(* IEC 61131-3 sources: Caravan/Archiv/12-04-19/Stations/MachineControl/MachineControl/Network/LseEasyMain, 1 file *)

(* ---- ONE_LseEasyMain_Table.st ---- *)
#define OBJECTS_CONFIG

#include "..\..\Source\Common\hmi_nuc.h"

FUNCTION GLOBAL TAB ONE_LseEasyMain
-1$UINT, 0$UINT,
0$UINT, 0$UINT,

40$UDINT,
TO_UDINT(3253426089), "HmiAsciiBuffer", 0$UINT, 0$UINT, 4$UINT,
TO_UDINT(3735923847), "HmiBaseList", 0$UINT, 0$UINT, 0$UINT,
TO_UDINT(2189921946), "HmiCanSendReceive", 0$UINT, 2$UINT, 1$UINT,
TO_UDINT(3930770040), "HmiChkBitList", 0$UINT, 2$UINT, 1$UINT,
TO_UDINT(845038353), "HmiColorMap", 0$UINT, 0$UINT, 1$UINT,
TO_UDINT(136722037), "HmiComPort", 0$UINT, 15$UINT, 0$UINT,
TO_UDINT(4239410787), "HmiComPortCan", 0$UINT, 14$UINT, 1$UINT,
TO_UDINT(2548286290), "HmiFile", 0$UINT, 4$UINT, 2$UINT,
TO_UDINT(1363967167), "HmiFont35", 0$UINT, 1$UINT, 1$UINT,
TO_UDINT(3893392983), "HmiFontList", 0$UINT, 3$UINT, 1$UINT,
TO_UDINT(3842677476), "HmiFunctionList", 0$UINT, 2$UINT, 1$UINT,
TO_UDINT(3385399892), "HmiFunctionList35", 0$UINT, 3$UINT, 1$UINT,
TO_UDINT(2724513001), "HmiImage35", 0$UINT, 3$UINT, 1$UINT,
TO_UDINT(3242935315), "HmiImageList", 0$UINT, 3$UINT, 1$UINT,
TO_UDINT(896341175), "HmiMapFile", 0$UINT, 0$UINT, 1$UINT,
TO_UDINT(3426238687), "HmiMemCircle", 0$UINT, 0$UINT, 1$UINT,
TO_UDINT(4250916264), "HmiMemImage", 0$UINT, 0$UINT, 1$UINT,
TO_UDINT(568511237), "HmiMemIO", 0$UINT, 0$UINT, 1$UINT,
TO_UDINT(1795655540), "HmiMemLine", 0$UINT, 0$UINT, 1$UINT,
TO_UDINT(2462046095), "HmiMemRectangle", 0$UINT, 0$UINT, 1$UINT,
TO_UDINT(2174260293), "HmiMemText", 0$UINT, 0$UINT, 1$UINT,
TO_UDINT(822070823), "HmiMemZorder", 0$UINT, 0$UINT, 1$UINT,
TO_UDINT(2613567777), "HmiProject35", 0$UINT, 4$UINT, 1$UINT,
TO_UDINT(2305619121), "HmiProjectList", 0$UINT, 1$UINT, 1$UINT,
TO_UDINT(2118014258), "HmiScreen", 0$UINT, 1$UINT, 1$UINT,
TO_UDINT(4172848962), "HmiSetUpList", 0$UINT, 2$UINT, 1$UINT,
TO_UDINT(1107224582), "HmiSetupList35", 0$UINT, 2$UINT, 1$UINT,
TO_UDINT(3851519469), "HmiShemeList", 0$UINT, 3$UINT, 4$UINT,
TO_UDINT(2500045939), "HmiShemeList35", 0$UINT, 3$UINT, 1$UINT,
TO_UDINT(4141094888), "HmiStateBit35", 0$UINT, 4$UINT, 1$UINT,
TO_UDINT(103556616), "HmiStrLib", 0$UINT, 2$UINT, 1$UINT,
TO_UDINT(2809265865), "HmiTextList", 0$UINT, 3$UINT, 1$UINT,
TO_UDINT(2738661249), "HmiTextList35", 0$UINT, 1$UINT, 1$UINT,
TO_UDINT(2548567416), "HmiUniBuffer", 0$UINT, 0$UINT, 10$UINT,
TO_UDINT(2706799507), "HmiUnitList", 0$UINT, 2$UINT, 1$UINT,
TO_UDINT(4154992490), "HmiUtils", 0$UINT, 2$UINT, 1$UINT,
TO_UDINT(1002095878), "HmiVarInfoList", 0$UINT, 1$UINT, 1$UINT,
TO_UDINT(3793961451), "HmiVarList", 0$UINT, 15$UINT, 1$UINT,
TO_UDINT(1599081198), "HmiVarList35", 0$UINT, 4$UINT, 1$UINT,
TO_UDINT(1518191916), "LseEasy", 1$UINT, 26$UINT, 1$UINT,

1$UINT, TO_UDINT(1344493304), "LSEEASY\HMICHKBITLIST\LABEL",
1$UINT, TO_UDINT(787249025), "LSEEASY\HMIFONTLIST\LABEL",
1$UINT, TO_UDINT(2117594790), "LSEEASY\HMIIMAGELIST\LABEL",
1$UINT, TO_UDINT(3002767849), "LSEEASY\HMIVARLIST\LABEL",

1$UINT, TO_UDINT(4084571679), "HMICOMPORTCAN1\CANSEND",

1$UINT, TO_UDINT(4275455085), "LSEEASY\HMICHKBITLIST",

1$UINT, TO_UDINT(846459028), "LSEEASY\HMICOLORMAP",

_NO_ATTR, TO_UDINT(1469804307), "HMICOMPORTCAN1",

1$UINT, TO_UDINT(1873895348), "HMICOMPORTCAN1\_BASE\FILE",
1$UINT, TO_UDINT(4182786947), "LSEEASY\FILE",

1$UINT, TO_UDINT(3760648512), "LSEEASY\HMIFONT35",

1$UINT, TO_UDINT(3896362450), "LSEEASY\HMIFONTLIST",

1$UINT, TO_UDINT(3636446795), "LSEEASY\HMIFUNCTIONLIST",

1$UINT, TO_UDINT(2190187032), "LSEEASY\HMIFUNCTIONLIST35",

1$UINT, TO_UDINT(2413249001), "LSEEASY\HMIIMAGE35",

1$UINT, TO_UDINT(1553538575), "LSEEASY\HMIIMAGELIST",

1$UINT, TO_UDINT(417239479), "LSEEASY\HMIMAPFILE",

1$UINT, TO_UDINT(2012497378), "LSEEASY\HMISCREEN\MEMCIRCLE",

1$UINT, TO_UDINT(975039261), "LSEEASY\HMISCREEN\MEMIMAGE",

1$UINT, TO_UDINT(3016924028), "LSEEASY\HMISCREEN\MEMIO",

1$UINT, TO_UDINT(4270949903), "LSEEASY\HMISCREEN\MEMLINE",

1$UINT, TO_UDINT(1370086185), "LSEEASY\HMISCREEN\MEMRECTANGLE",

1$UINT, TO_UDINT(336500030), "LSEEASY\HMISCREEN\MEMTEXT",

1$UINT, TO_UDINT(2335427354), "LSEEASY\HMISCREEN\MEMZORDER",

1$UINT, TO_UDINT(102087485), "LSEEASY\HMIPROJECT35",

1$UINT, TO_UDINT(3836054740), "LSEEASY\HMIPROJECTLIST",

1$UINT, TO_UDINT(3478444237), "LSEEASY\HMISCREEN",

1$UINT, TO_UDINT(1701496158), "LSEEASY\HMISETUPLIST",

1$UINT, TO_UDINT(741838947), "LSEEASY\HMISETUPLIST35",

1$UINT, TO_UDINT(2459869223), "LSEEASY\HMIFONTSHEMELIST",
1$UINT, TO_UDINT(1282849623), "LSEEASY\HMIIMAGESHEMELIST",
1$UINT, TO_UDINT(3937490271), "LSEEASY\HMITEXTSHEMELIST",
1$UINT, TO_UDINT(3509062318), "LSEEASY\HMIVARLIST\HMIUNITSHEMELIST",

1$UINT, TO_UDINT(4174042134), "LSEEASY\HMISHEMELIST35",

1$UINT, TO_UDINT(3796408829), "LSEEASY\HMISTATEBIT35",

1$UINT, TO_UDINT(1881447452), "LSEEASY\STRINGLIB",

1$UINT, TO_UDINT(2807844172), "LSEEASY\HMITEXTLIST",

1$UINT, TO_UDINT(3080726932), "LSEEASY\HMITEXTLIST35",

1$UINT, TO_UDINT(2308124733), "LSEEASY\HMITEXTLIST\TEXTLIST00",
1$UINT, TO_UDINT(4271112363), "LSEEASY\HMITEXTLIST\TEXTLIST01",
1$UINT, TO_UDINT(1738363153), "LSEEASY\HMITEXTLIST\TEXTLIST02",
1$UINT, TO_UDINT(278552967), "LSEEASY\HMITEXTLIST\TEXTLIST03",
1$UINT, TO_UDINT(2399073316), "LSEEASY\HMITEXTLIST\TEXTLIST04",
1$UINT, TO_UDINT(4193895602), "LSEEASY\HMITEXTLIST\TEXTLIST05",
1$UINT, TO_UDINT(1626379528), "LSEEASY\HMITEXTLIST\TEXTLIST06",
1$UINT, TO_UDINT(402105758), "LSEEASY\HMITEXTLIST\TEXTLIST07",
1$UINT, TO_UDINT(2269689871), "LSEEASY\HMITEXTLIST\TEXTLIST08",
1$UINT, TO_UDINT(4031744153), "LSEEASY\HMITEXTLIST\TEXTLIST09",

1$UINT, TO_UDINT(200861884), "LSEEASY\HMIVARLIST\UNITINFO",

1$UINT, TO_UDINT(2530016337), "LSEEASY\HMIUTILS",

1$UINT, TO_UDINT(3991554070), "LSEEASY\HMIVARLIST\VARINFO",

1$UINT, TO_UDINT(3482371307), "LSEEASY\HMIVARLIST",

1$UINT, TO_UDINT(3263320306), "LSEEASY\HMIVARLIST35",

_NO_ATTR, TO_UDINT(1518191916), "LSEEASY",

//Internal connections
0$UDINT,
52$UDINT,
TO_UDINT(5), "Label", TO_UDINT(0),
TO_UDINT(7), "File", TO_UDINT(8),
TO_UDINT(7), "CanSend", TO_UDINT(4),
TO_UDINT(11), "Label", TO_UDINT(1),
TO_UDINT(15), "Label", TO_UDINT(2),
TO_UDINT(26), "MemRectangle", TO_UDINT(21),
TO_UDINT(26), "MemText", TO_UDINT(22),
TO_UDINT(26), "MemIO", TO_UDINT(19),
TO_UDINT(26), "MemCircle", TO_UDINT(17),
TO_UDINT(26), "MemLine", TO_UDINT(20),
TO_UDINT(26), "MemImage", TO_UDINT(18),
TO_UDINT(26), "MemZorder", TO_UDINT(23),
TO_UDINT(36), "TextList00", TO_UDINT(38),
TO_UDINT(36), "TextList01", TO_UDINT(39),
TO_UDINT(36), "TextList02", TO_UDINT(40),
TO_UDINT(36), "TextList03", TO_UDINT(41),
TO_UDINT(36), "TextList04", TO_UDINT(42),
TO_UDINT(36), "TextList05", TO_UDINT(43),
TO_UDINT(36), "TextList06", TO_UDINT(44),
TO_UDINT(36), "TextList07", TO_UDINT(45),
TO_UDINT(36), "TextList08", TO_UDINT(46),
TO_UDINT(36), "TextList09", TO_UDINT(47),
TO_UDINT(51), "UnitInfo", TO_UDINT(48),
TO_UDINT(51), "Label", TO_UDINT(3),
TO_UDINT(51), "VarInfo", TO_UDINT(50),
TO_UDINT(51), "HmiUnitShemeList", TO_UDINT(32),
TO_UDINT(53), "HmiImageList", TO_UDINT(15),
TO_UDINT(53), "HmiFunctionList", TO_UDINT(12),
TO_UDINT(53), "HmiScreen", TO_UDINT(26),
TO_UDINT(53), "HmiFontList", TO_UDINT(11),
TO_UDINT(53), "HmiVarList", TO_UDINT(51),
TO_UDINT(53), "HmiColorMap", TO_UDINT(6),
TO_UDINT(53), "HmiProjectList", TO_UDINT(25),
TO_UDINT(53), "HmiProject35", TO_UDINT(24),
TO_UDINT(53), "HmiTextList", TO_UDINT(36),
TO_UDINT(53), "HmiVarList35", TO_UDINT(52),
TO_UDINT(53), "HmiFont35", TO_UDINT(10),
TO_UDINT(53), "HmiImage35", TO_UDINT(14),
TO_UDINT(53), "HmiSetUpList", TO_UDINT(27),
TO_UDINT(53), "HmiFunctionList35", TO_UDINT(13),
TO_UDINT(53), "HmiShemeList35", TO_UDINT(33),
TO_UDINT(53), "HmiFontShemeList", TO_UDINT(29),
TO_UDINT(53), "HmiTextShemeList", TO_UDINT(31),
TO_UDINT(53), "HmiImageShemeList", TO_UDINT(30),
TO_UDINT(53), "HmiSetupList35", TO_UDINT(28),
TO_UDINT(53), "StringLib", TO_UDINT(35),
TO_UDINT(53), "File", TO_UDINT(9),
TO_UDINT(53), "HmiUtils", TO_UDINT(49),
TO_UDINT(53), "HmiTextList35", TO_UDINT(37),
TO_UDINT(53), "HmiChkBitList", TO_UDINT(5),
TO_UDINT(53), "HmiStateBit35", TO_UDINT(34),
TO_UDINT(53), "HmiMapFile", TO_UDINT(16),
0$UDINT,
33$UDINT,
TO_UDINT(5), "File", TO_UDINT(9), "ClassSvr",
TO_UDINT(5), "VarList", TO_UDINT(51), "ClassSvr",
TO_UDINT(5), "StringLib", TO_UDINT(35), "ClassSvr",
TO_UDINT(6), "File", TO_UDINT(9), "ClassSvr",
TO_UDINT(11), "File", TO_UDINT(9), "ClassSvr",
TO_UDINT(11), "StringLib", TO_UDINT(35), "ClassSvr",
TO_UDINT(12), "File", TO_UDINT(9), "ClassSvr",
TO_UDINT(13), "HmiVarList", TO_UDINT(51), "ClassSvr",
TO_UDINT(15), "File", TO_UDINT(9), "ClassSvr",
TO_UDINT(15), "StringLib", TO_UDINT(35), "ClassSvr",
TO_UDINT(16), "File", TO_UDINT(9), "ClassSvr",
TO_UDINT(16), "VarList", TO_UDINT(51), "ClassSvr",
TO_UDINT(16), "StateBit", TO_UDINT(34), "ClassSvr",
TO_UDINT(16), "StringLib", TO_UDINT(35), "ClassSvr",
TO_UDINT(25), "File", TO_UDINT(9), "ClassSvr",
TO_UDINT(25), "StringLib", TO_UDINT(35), "ClassSvr",
TO_UDINT(26), "File", TO_UDINT(9), "ClassSvr",
TO_UDINT(27), "File", TO_UDINT(9), "ClassSvr",
TO_UDINT(29), "File", TO_UDINT(9), "ClassSvr",
TO_UDINT(30), "File", TO_UDINT(9), "ClassSvr",
TO_UDINT(31), "File", TO_UDINT(9), "ClassSvr",
TO_UDINT(34), "ChkBit", TO_UDINT(5), "ClassSvr",
TO_UDINT(34), "VarList", TO_UDINT(51), "ClassSvr",
TO_UDINT(34), "StringLib", TO_UDINT(35), "ClassSvr",
TO_UDINT(36), "File", TO_UDINT(9), "ClassSvr",
TO_UDINT(36), "StringLib", TO_UDINT(35), "ClassSvr",
TO_UDINT(36), "HmiVarList", TO_UDINT(51), "ClassSvr",
TO_UDINT(36), "HmiTextList35", TO_UDINT(37), "ClassSvr",
TO_UDINT(51), "File", TO_UDINT(9), "ClassSvr",
TO_UDINT(51), "StringLib", TO_UDINT(35), "ClassSvr",
TO_UDINT(51), "TextList", TO_UDINT(36), "ClassSvr",
TO_UDINT(51), "HmiVarList35", TO_UDINT(52), "ClassSvr",
TO_UDINT(53), "ComPort", TO_UDINT(7), "ClassSvr",

//Initialization values
0$UDINT,
17$UDINT,
TO_UDINT(4), "CanNodeDisplay", TO_UDINT(1),//|LseEasyMain.HmiComPortCan1\CanSend.CanNodeDisplay;
TO_UDINT(4), "CanInterface", TO_UDINT(1),//|LseEasyMain.HmiComPortCan1\CanSend.CanInterface;
TO_UDINT(4), "CanRxMsgID", TO_UDINT(16#40),//|LseEasyMain.HmiComPortCan1\CanSend.CanRxMsgID;
TO_UDINT(4), "CanTxMsgID", TO_UDINT(16#20),//|LseEasyMain.HmiComPortCan1\CanSend.CanTxMsgID;
TO_UDINT(7), "CanNodeDisplay", TO_UDINT(1),//|LseEasyMain.HmiComPortCan1.CanNodeDisplay;
TO_UDINT(7), "CanInterface", TO_UDINT(1),//|LseEasyMain.HmiComPortCan1.CanInterface;
TO_UDINT(7), "CanRxMsgID", TO_UDINT(16#40),//|LseEasyMain.HmiComPortCan1.CanRxMsgID;
TO_UDINT(7), "CanTxMsgID", TO_UDINT(16#20),//|LseEasyMain.HmiComPortCan1.CanTxMsgID;
TO_UDINT(34), "ComPort", TO_UDINT(0),//|LseEasyMain.LseEasy\HmiStateBit35.ComPort;
TO_UDINT(51), "ComPort", TO_UDINT(0),//|LseEasyMain.LseEasy\HmiVarList.ComPort;
TO_UDINT(53), "ActLanguage", TO_UDINT(0),//|LseEasyMain.LseEasy.ActLanguage;
TO_UDINT(53), "ComPort", TO_UDINT(0),//|LseEasyMain.LseEasy.ComPort;
TO_UDINT(53), "ProjectPath", TO_UDINT(0),//|LseEasyMain.LseEasy.ProjectPath;
TO_UDINT(53), "TempInterval", TO_UDINT(1000),//|LseEasyMain.LseEasy.TempInterval;
TO_UDINT(53), "BackLightOff", TO_UDINT(10000),//|LseEasyMain.LseEasy.BackLightOff;
TO_UDINT(53), "OverloadLight", TO_UDINT(-1),//|LseEasyMain.LseEasy.OverloadLight;
TO_UDINT(53), "AutoFirmwareUpdate", TO_UDINT(0),//|LseEasyMain.LseEasy.AutoFirmwareUpdate;

//Symbolic initialization values
0$UDINT,
0$UDINT,

//Initialization of string values
0$UDINT,
0$UDINT,

//Configuration of tasks (RealTime, Cyclic, Background)
0$UDINT,
0$UDINT,

0$UDINT,
0$UDINT,

0$UDINT,
1$UDINT,
TO_UDINT(53), (-1)$UDINT, 4194303$DINT, 	//LSEEASY

//External connections
0$UDINT,
0$UDINT,

//Magic internal connections
0$UDINT,
45$UDINT,
TO_UDINT(0), "File", TO_UDINT(5), "File",
TO_UDINT(0), "StringLib", TO_UDINT(5), "StringLib",
TO_UDINT(1), "File", TO_UDINT(11), "File",
TO_UDINT(1), "StringLib", TO_UDINT(11), "StringLib",
TO_UDINT(2), "File", TO_UDINT(15), "File",
TO_UDINT(2), "StringLib", TO_UDINT(15), "StringLib",
TO_UDINT(51), "ComPort", TO_UDINT(53), "ComPort",
TO_UDINT(3), "File", TO_UDINT(51), "File",
TO_UDINT(3), "StringLib", TO_UDINT(51), "StringLib",
TO_UDINT(4), "CanNodeDisplay", TO_UDINT(7), "CanNodeDisplay",
TO_UDINT(4), "CanInterface", TO_UDINT(7), "CanInterface",
TO_UDINT(4), "CanRxMsgID", TO_UDINT(7), "CanRxMsgID",
TO_UDINT(4), "CanTxMsgID", TO_UDINT(7), "CanTxMsgID",
TO_UDINT(4), "CoCanLib", TO_UDINT(7), "CoCanLib",
TO_UDINT(17), "File", TO_UDINT(26), "File",
TO_UDINT(18), "File", TO_UDINT(26), "File",
TO_UDINT(19), "File", TO_UDINT(26), "File",
TO_UDINT(20), "File", TO_UDINT(26), "File",
TO_UDINT(21), "File", TO_UDINT(26), "File",
TO_UDINT(22), "File", TO_UDINT(26), "File",
TO_UDINT(23), "File", TO_UDINT(26), "File",
TO_UDINT(32), "File", TO_UDINT(51), "File",
TO_UDINT(34), "ComPort", TO_UDINT(53), "ComPort",
TO_UDINT(38), "File", TO_UDINT(36), "File",
TO_UDINT(38), "StringLib", TO_UDINT(36), "StringLib",
TO_UDINT(39), "File", TO_UDINT(36), "File",
TO_UDINT(39), "StringLib", TO_UDINT(36), "StringLib",
TO_UDINT(40), "File", TO_UDINT(36), "File",
TO_UDINT(40), "StringLib", TO_UDINT(36), "StringLib",
TO_UDINT(41), "File", TO_UDINT(36), "File",
TO_UDINT(41), "StringLib", TO_UDINT(36), "StringLib",
TO_UDINT(42), "File", TO_UDINT(36), "File",
TO_UDINT(42), "StringLib", TO_UDINT(36), "StringLib",
TO_UDINT(43), "File", TO_UDINT(36), "File",
TO_UDINT(43), "StringLib", TO_UDINT(36), "StringLib",
TO_UDINT(44), "File", TO_UDINT(36), "File",
TO_UDINT(44), "StringLib", TO_UDINT(36), "StringLib",
TO_UDINT(45), "File", TO_UDINT(36), "File",
TO_UDINT(45), "StringLib", TO_UDINT(36), "StringLib",
TO_UDINT(46), "File", TO_UDINT(36), "File",
TO_UDINT(46), "StringLib", TO_UDINT(36), "StringLib",
TO_UDINT(47), "File", TO_UDINT(36), "File",
TO_UDINT(47), "StringLib", TO_UDINT(36), "StringLib",
TO_UDINT(48), "File", TO_UDINT(51), "File",
TO_UDINT(50), "File", TO_UDINT(51), "File",

//Configuration of timeslots of tasks (RealTime, Cyclic)
#ifdef __LSLLDR_TIMESLOTS__
0$UDINT,
0$UDINT,

0$UDINT,
0$UDINT,

#endif //__LSLLDR_TIMESLOTS__

//MultiMaster connections
#ifdef __LSLLDR_MULTIMASTER__
0$UDINT,
0$UDINT,
#endif //__LSLLDR_MULTIMASTER__

//Configuration for task ID (RealTime, CyclicTime)
#ifdef __LSLLDR_TASKID__
"\\\\TASKS2  "
0$UDINT,
0$UDINT,

0$UDINT,
0$UDINT,

0$UDINT,
1$UDINT,
(0)$UDINT, 	//LSEEASY

#endif //__LSLLDR_TASKID__

END_FUNCTION
